Staubli VAL3: HMI_IO.pjx

--- HMI_IO.pjx ---
Parameters version=s8.10.3Cs9_BS2093 stackSize=5000 millimeterUnit=true
Program file=bind.pgx
Program file=comment.pgx
Program file=getSize.pgx
Program file=init.pgx
Program file=IOcomment.pgx
Program file=main.pgx
Program file=SetbtnColor.pgx
Program file=setCount.pgx
Program file=setIOStatus.pgx
Program file=setIOvisible.pgx
Program file=setLabelValue.pgx
Program file=setPage.pgx
Program file=start.pgx
Program file=stop.pgx
Data file=HMI_IO.dtx
Library alias=util path=Disk://HMI_cs9/HMI_util/HMI_util.pjx
Library alias=rs path=Disk://source/projectSource/robotStatus/robotStatus.pjx
Library alias=io path=Disk://source/projectSource/io/io.pjx

--- HMI_IO.dtx ---
mdesc mNomSpeed
num nPage
num nPageIndex
num nItemIndex
public bool bBool[11]
public string sUsingBus
bool bComment[16]
public string sLabel[16]
num nShowPageIndex
string sShowPageIndex
string sPageNum
public string sComment[16]
num nType
num nSelType
bool bRefresh
public string sValue[16]
bool bBtnHidden
bool bLabelHidden
num _nClock
bool bBack
num nDigCount
num nAngCount
bool bConfirm
bool bCancel

--- main.pgx ---
public program main()
  local bool l_bExit
  local bool l_bResult
begin
  do
    if util:sPage!="IO"
      util:sPage="IO"
      call util:loadingPage()
      call bind()
      call init()
      userPage(util:sPage)
      delay(0.5)
      bRefresh=true
    endIf
    //btn click
    if bBool[1]
      bBool[1]=false
      nSelType=0
      bRefresh=true
      call SetbtnColor(nSelType)
      //din
    elseIf bBool[2]
      bBool[2]=false
      nSelType=1
      bRefresh=true
      call SetbtnColor(nSelType)
      //dout
    elseIf bBool[3]
      bBool[3]=false
      nSelType=2
      bRefresh=true
      call SetbtnColor(nSelType)
      //ain
    elseIf bBool[4]
      bBool[4]=false
      nSelType=3
      bRefresh=true
      call SetbtnColor(nSelType)
      //dout
    elseIf bBool[5]
      bBool[5]=false
      //change bus
      l_bResult=userPageConfirm("是否切换到总线协议："+sUsingBus)
      if l_bResult
        call io:linkIO(sUsingBus)
        rs:sBusUsing=sUsingBus
        rs:libSave()
        delay(0.1)
        userPageAlert("通讯协议已切换到"+rs:sBusUsing+"重启app生效")
      endIf
    elseIf bBool[6]
      bBool[6]=false
      //head page
      nPageIndex=0
      bRefresh=true
    elseIf bBool[7]
      bBool[7]=false
      //backward
      if nPageIndex>0
        nPageIndex=nPageIndex-1
      else
        nPageIndex=0
      endIf
      bRefresh=true
    elseIf bBool[8]
      bBool[8]=false
      //forward
      if nPageIndex<nPage-1
        nPageIndex=nPageIndex+1
      else
        nPageIndex=nPage-1
      endIf
      bRefresh=true
    elseIf bBool[9]
      bBool[9]=false
      //end page
      nPageIndex=nPage-1
      bRefresh=true
    elseIf bBool[10]
      bBool[10]=false
      call setCount()
    elseIf bBack==true
      bBack=false
      l_bExit=true
    endIf
    call comment(bRefresh)
    //refresh
    if bRefresh
      bRefresh=false
      call setPage(nSelType)
      call setLabelValue(nSelType)
      call setIOvisible(nSelType)
      delay(0)
    endIf
    if clock()-_nClock>0.1
      call setIOStatus(nSelType)
      _nClock=clock()
    endIf
    delay(0.1)
  until l_bExit==true
end

--- start.pgx ---
program start()
begin
end

--- bind.pgx ---
public program bind()
  local string l_sbtn
  local string l_slbl
  local num l_i
begin
  //btn bind
  for l_i = 1 to 10 step 1
    l_sbtn="btn"+toString("",l_i)
    bBool[l_i]=false
    userPageBindClick("IO",l_sbtn,bBool[l_i],true)
  endFor
  userPageBindClick("IO","btnback",bBack,true)
  //label bind
  userPageBind("IO","lblpageIndex","innerHTML",sShowPageIndex,1,"r")
  userPageBind("IO","lblpage","innerHTML",sPageNum,1,"r")
  //label Click
  for l_i = 0 to 15
    l_slbl="lbl"+toString("",20+l_i)
    //comment
    userPageBindClick("IO",l_slbl,bComment[l_i],true)
  endFor
  //innerHTML
  for l_i = 0 to 15
    l_slbl="lbl"+toString("",l_i)
    //title
    userPageBind("IO",l_slbl,"innerHTML",sLabel[l_i],1,"r")
  endFor
  for l_i = 0 to 15
    l_slbl="lbl"+toString("",40+l_i)
    //aio value
    userPageBind("IO",l_slbl,"innerHTML",sValue[l_i],1,"r")
  endFor
  for l_i = 0 to 15
    l_slbl="lbl"+toString("",20+l_i)
    //comment
    userPageBind("IO",l_slbl,"innerHTML",sComment[l_i],1,"r")
  endFor

  //combox
  userPageBind("IO","cbx1","value",sUsingBus,1,"rw")

end

--- comment.pgx ---
public program comment(bool& x_bRefresh)
  local string l_sString
  local bool l_bResult
  local num l_i
  local num l_nIndex
begin
  for l_i = 0 to size(bComment)-1
    if bComment[l_i]
      bComment[l_i]=false
      l_bResult=userPagePrompt("注释：",l_sString)
      if l_bResult
        l_nIndex=nPageIndex*16+l_i
        //Modify by Liu Zhengang 20251103
        switch nSelType
          case 0,1
            if 15<l_nIndex and l_nIndex<96
              call IOcomment(nSelType,l_nIndex,l_sString)
            else
              userPageAlert("此信号不可修改注释！")
            endIf
            io:libSave()
            delay(0.1)
            x_bRefresh=true
          break
          case 2,3
            if 4<l_nIndex and l_nIndex<20
              call IOcomment(nSelType,l_nIndex,l_sString)
            else
              userPageAlert("此信号不可修改注释！")
            endIf
            io:libSave()
            delay(0.1)
            x_bRefresh=true
          break
        endSwitch
      endIf
    endIf
  endFor
end

--- getSize.pgx ---
public program getSize(num& x_nSize, num& x_nSize1)
begin
  if io:nMaxdigital%16!=0 and nPageIndex==nPage-1
    x_nSize=io:nMaxdigital%16
  else
    x_nSize=16
  endIf
 if io:nMaxAnalog%16!=0 and nPageIndex==nPage-1
    x_nSize1=io:nMaxAnalog%16
  else
    x_nSize1=16
  endIf
end

--- init.pgx ---
public program init()
  local num l_i
begin
  nPage=0
  nPageIndex=0
  nItemIndex=0

  nPage=roundUp(size(io:dInItem)/16)
  sShowPageIndex=toString("",nPageIndex+1)
  sPageNum=toString("",nPage)
  sUsingBus=rs:sBusUsing
  nSelType=0
  call SetbtnColor(nSelType)
  for l_i = 0 to 15
    sLabel[l_i]=""
    sComment[l_i]=""
  endFor
  if io:nMaxAnalog<=0
    userPageSet("IO","btn3","disabled",true)
    userPageSet("IO","btn4","disabled",true)
    popUpMsg("模拟量数量未设置")
  endIf
  //  //list
  //  for l_i = 0 to 15
  //    sLabel[l_i]="dIn["+toString("",l_i+16*nPageIndex)+"]"
  //    sComment[l_i]=io:dInItem[l_i+16*nPageIndex].sComment
  //  endFor

end

--- IOcomment.pgx ---
public program IOcomment(num x_nType, num x_nIndex, string x_sComment)
begin
  switch x_nType
    case 0
      io:dInItem[x_nIndex].sComment=x_sComment
      io:sCommentDin[x_nIndex]=x_sComment
    break
    case 1
      io:dOutItem[x_nIndex].sComment=x_sComment
      io:sCommentDout[x_nIndex]=x_sComment
    break
    case 2
      io:aInItem[x_nIndex].sComment=x_sComment
      io:sCommentAin[x_nIndex]=x_sComment
    break
    case 3
      io:aOutItem[x_nIndex].sComment=x_sComment
      io:sCommentAout[x_nIndex]=x_sComment
    break

  endSwitch

  io:libSave()
  delay(0)
end

--- SetbtnColor.pgx ---
public program SetbtnColor(num x_nNum)
  local string l_selColor
  local string l_sNULLcolor
begin
  l_selColor="#9999FF"
  l_sNULLcolor="#FFFFFF"
  switch x_nNum
    case 0
      userPageSet("IO","btn1","style.backgroundColor",l_selColor)
      userPageSet("IO","btn2","style.backgroundColor",l_sNULLcolor)
      userPageSet("IO","btn3","style.backgroundColor",l_sNULLcolor)
      userPageSet("IO","btn4","style.backgroundColor",l_sNULLcolor)
    break
    case 1
      userPageSet("IO","btn1","style.backgroundColor",l_sNULLcolor)
      userPageSet("IO","btn2","style.backgroundColor",l_selColor)
      userPageSet("IO","btn3","style.backgroundColor",l_sNULLcolor)
      userPageSet("IO","btn4","style.backgroundColor",l_sNULLcolor)
    break
    case 2
      userPageSet("IO","btn1","style.backgroundColor",l_sNULLcolor)
      userPageSet("IO","btn2","style.backgroundColor",l_sNULLcolor)
      userPageSet("IO","btn3","style.backgroundColor",l_selColor)
      userPageSet("IO","btn4","style.backgroundColor",l_sNULLcolor)
    break
    case 3
      userPageSet("IO","btn1","style.backgroundColor",l_sNULLcolor)
      userPageSet("IO","btn2","style.backgroundColor",l_sNULLcolor)
      userPageSet("IO","btn3","style.backgroundColor",l_sNULLcolor)
      userPageSet("IO","btn4","style.backgroundColor",l_selColor)
    break
  endSwitch
end

--- setCount.pgx ---
public program setCount()
  local num l_nSize1
  local num l_nSize2
  local bool l_bExit
begin
  do
    if util:sPage!="setCount"
      util:sPage="setCount"
      nDigCount=io:nMaxdigital
      nAngCount=io:nMaxAnalog
      userPageBind("setCount","nmb1","value",nDigCount,1,"rw")
      userPageBind("setCount","nmb2","value",nAngCount,1,"rw")
      userPageBindClick("setCount","btn1",bConfirm,true)
      userPageBindClick("setCount","btn2",bCancel,true)
      userPage(util:sPage)
      delay(0.5)
    endIf


    //btn
    if bConfirm
      bConfirm=false
      call io:getAngIOSize(l_nSize1)
      call io:getDigIOSize(l_nSize2)
      io:nMaxdigital=nDigCount
      io:nMaxAnalog=nAngCount
      call io:linkIO(rs:sBusUsing)
      io:libSave()
      popUpMsg("IO数据长度已更新")
      delay(0.5)
      l_bExit=true
    elseIf bCancel
      bCancel=false

      l_bExit=true

    endIf

    delay(0)
  until l_bExit==true
end

--- setIOStatus.pgx ---
public program setIOStatus(num x_nType)
  local num l_nSize
  local string l_selColor
  local string l_sNullColor
  local string l_sbtn
  local string l_sErrColor
  local string l_slabel
  local num l_nValue
  local num l_i
  local num l_nSize1
  local string l_slbl1
  local string l_slbl2
begin
  l_selColor="#33FF33"
  l_sNullColor="#FFFFFF"
  l_sErrColor="#C8C8C8"
  call getSize(l_nSize,l_nSize1)
  //  if l_nSize<16
  //    for l_i = l_nSize to 15
  //      l_sbtn="btn"+toString("",60+l_i)
  //      l_slbl1="lbl"+toString("",20+l_i)
  //      l_slbl2="lbl"+toString("",l_i)
  //      userPageSet("IO",l_sbtn,"style.visibility","hidden")
  //      userPageSet("IO",l_slbl1,"style.visibility","hidden")
  //      userPageSet("IO",l_slbl2,"style.visibility","hidden")
  //    endFor
  //  endIf
  //  if l_nSize1<16
  //    for l_i = l_nSize1 to 15
  //      l_sbtn="lbl"+toString("",40+l_i)
  //      l_slbl1="lbl"+toString("",20+l_i)
  //      l_slbl2="lbl"+toString("",l_i)
  //      userPageSet("IO",l_sbtn,"style.visibility","hidden")
  //      userPageSet("IO",l_slbl1,"style.visibility","hidden")
  //      userPageSet("IO",l_slbl2,"style.visibility","hidden")
  //    endFor
  //  endIf

  switch x_nType
    case 0
      for l_i = 0 to l_nSize-1
        l_sbtn="btn"+toString("",60+l_i)
        //     userPageSet("IO",l_sbtn,"style.visibility","visible")
        if ioStatus(io:dInItem[l_i+nPageIndex*16].dDio)>-1
          l_nValue=dioGet(io:dInItem[l_i+nPageIndex*16].dDio)
          if l_nValue==1
            userPageSet("IO",l_sbtn,"style.backgroundColor",l_selColor)
          else
            userPageSet("IO",l_sbtn,"style.backgroundColor",l_sNullColor)
          endIf
        else
          userPageSet("IO",l_sbtn,"style.backgroundColor",l_sErrColor)
        endIf
      endFor
    break
    case 1
      for l_i = 0 to l_nSize-1
        l_sbtn="btn"+toString("",60+l_i)
        //     userPageSet("IO",l_sbtn,"style.visibility","visible")
        if ioStatus(io:dOutItem[l_i+nPageIndex*16].dDio)>-1
          l_nValue=dioGet(io:dOutItem[l_i+nPageIndex*16].dDio)
          if l_nValue==1
            userPageSet("IO",l_sbtn,"style.backgroundColor",l_selColor)
          else
            userPageSet("IO",l_sbtn,"style.backgroundColor",l_sNullColor)
          endIf
        else
          userPageSet("IO",l_sbtn,"style.backgroundColor",l_sErrColor)
        endIf
      endFor
    break
    case 2
      for l_i = 0 to l_nSize1-1
        l_slabel="lbl"+toString("",40+l_i)
        //       userPageSet("IO",l_slabel,"style.visibility","visible")
        if ioStatus(io:aInItem[l_i+nPageIndex*16].aAio)>-1
          l_nValue=aioGet(io:aInItem[l_i+nPageIndex*16].aAio)
          sValue[l_i]=toString(".2",l_nValue)
        else
          sValue[l_i]="?"
        endIf
      endFor
    break
    case 3
      for l_i = 0 to l_nSize1-1
        l_slabel="lbl"+toString("",40+l_i)
        //      userPageSet("IO",l_slabel,"style.visibility","visible")
        if ioStatus(io:aOutItem[l_i+nPageIndex*16].aAio)>-1
          l_nValue=aioGet(io:aOutItem[l_i+nPageIndex*16].aAio)
          sValue[l_i]=toString(".2",l_nValue)
        else
          sValue[l_i]="?"
        endIf
      endFor
    break

  endSwitch

end

--- setIOvisible.pgx ---
public program setIOvisible(num x_nType)
  local string l_sbtn
  local num l_i
  local string l_slabel
  local num l_nSize
  local string l_slbl
  local string l_slbl1
  local string l_slbl2
  local num l_nSize1
begin
  call getSize(l_nSize,l_nSize1)
  switch x_nType
    case 0,1
      for l_i = 0 to 15
        l_slbl="lbl"+toString("",40+l_i)
        userPageSet("IO",l_slbl,"style.visibility","hidden")
      endFor
      for l_i = 0 to l_nSize-1
        l_slbl="lbl"+toString("",l_i)
        l_slbl1="lbl"+toString("",20+l_i)
        l_slbl2="btn"+toString("",60+l_i)
        userPageSet("IO",l_slbl,"style.visibility","visible")
        userPageSet("IO",l_slbl1,"style.visibility","visible")
        userPageSet("IO",l_slbl2,"style.visibility","visible")
      endFor
      if l_nSize<16
        for l_i = l_nSize to 15
          l_slbl="lbl"+toString("",l_i)
          l_slbl1="lbl"+toString("",20+l_i)
          l_slbl2="btn"+toString("",60+l_i)
          userPageSet("IO",l_slbl,"style.visibility","hidden")
          userPageSet("IO",l_slbl1,"style.visibility","hidden")
          userPageSet("IO",l_slbl2,"style.visibility","hidden")
        endFor
      endIf
    break
    case 2,3
      for l_i = 0 to 15
        l_slbl="btn"+toString("",60+l_i)
        userPageSet("IO",l_slbl,"style.visibility","hidden")
      endFor
      for l_i = 0 to l_nSize1-1
        l_slbl="lbl"+toString("",l_i)
        l_slbl1="lbl"+toString("",20+l_i)
        l_slbl2="lbl"+toString("",40+l_i)
        userPageSet("IO",l_slbl,"style.visibility","visible")
        userPageSet("IO",l_slbl1,"style.visibility","visible")
        userPageSet("IO",l_slbl2,"style.visibility","visible")
      endFor
      if l_nSize1<16
        for l_i = l_nSize1 to 15
          l_slbl="lbl"+toString("",l_i)
          l_slbl1="lbl"+toString("",20+l_i)
          l_slbl2="lbl"+toString("",40+l_i)
          userPageSet("IO",l_slbl,"style.visibility","hidden")
          userPageSet("IO",l_slbl1,"style.visibility","hidden")
          userPageSet("IO",l_slbl2,"style.visibility","hidden")
        endFor
      endIf
    break
  endSwitch
end

--- setLabelValue.pgx ---
public program setLabelValue(num x_nType)
  local num l_nSize
  local num l_i
  local string l_slabel
  local num l_nSize1
begin

  call getSize(l_nSize,l_nSize1)
  //
  switch x_nType
    case 0
      for l_i = 0 to l_nSize-1
        sLabel[l_i]=toString("",l_i+16*nPageIndex)+".dIn["+toString("",l_i+16*nPageIndex)+"]"
        sComment[l_i]=io:dInItem[l_i+16*nPageIndex].sComment
      endFor
    break
    case 1
      for l_i = 0 to l_nSize-1
        sLabel[l_i]=toString("",l_i+16*nPageIndex)+".dOut["+toString("",l_i+16*nPageIndex)+"]"
        sComment[l_i]=io:dOutItem[l_i+16*nPageIndex].sComment
      endFor
    break
    case 2
      for l_i = 0 to l_nSize1-1
        sLabel[l_i]=toString("",l_i+16*nPageIndex)+".aIn["+toString("",l_i+16*nPageIndex)+"]"
        sComment[l_i]=io:aInItem[l_i+16*nPageIndex].sComment
      endFor
    break
    case 3
      for l_i = 0 to l_nSize1-1
        sLabel[l_i]=toString("",l_i+16*nPageIndex)+".aOut["+toString("",l_i+16*nPageIndex)+"]"
        sComment[l_i]=io:aOutItem[l_i+16*nPageIndex].sComment
      endFor

    break
  endSwitch

end

--- setPage.pgx ---
public program setPage(num x_nType)
begin
  switch x_nType
    case 0,1

      nPage=roundUp(io:nMaxdigital/16)

    break
    case 2,3
      nPage=roundUp(io:nMaxAnalog/16)
      if nPageIndex>nPage-1
        nPageIndex=0
      endIf
    break
  endSwitch
  sPageNum=toString("",nPage)
  sShowPageIndex=toString("",nPageIndex+1)
end

--- stop.pgx ---
program stop()
begin
end
